FUNCTION_BLOCK FB_StartupReadiness_Tests EXTENDS TcUnit.FB_TestSuite

Power_To_Home_Handoff();
Abort_Cannot_Become_Online();
Error_And_Park_Win();
Completion_Requires_Operational();
Explicit_Abort_Invalidates_Completed_Startup();
Repeated_Start_Does_Not_Reset_Calibration();
Suspended_Automatic_Needs_New_Startup();
Start_While_Initialized_Restarts_Calibration();
Error_Needs_New_Startup();
Parking_Invalidates_Completed_Startup();
Preparation_Stays_0_7_Until_Calibrating();

METHOD PRIVATE Power_To_Home_Handoff
VAR
    fb : BROTLib.FB_StartupReadiness;
END_VAR
TEST('Power_To_Home_Handoff');
fb(Start := TRUE, Parked := TRUE);
AssertEquals_LREAL(0.7, fb.ReadyState, 0.0001, 'preparation, even if parked flag has not cleared');
fb(Start := FALSE, Calibrating := TRUE, Parked := FALSE, Operational := TRUE);
AssertEquals_LREAL(0.8, fb.ReadyState, 0.0001, 'calibration, axes mechanically ready');
fb(Calibrating := FALSE);
AssertEquals_LREAL(0.8, fb.ReadyState, 0.0001, 'handoff/intermediate standstill stays pending');
fb(Completed := TRUE);
AssertEquals_LREAL(1.0, fb.ReadyState, 0.0001, 'only terminal completion is online');
fb(Completed := FALSE);
AssertEquals_LREAL(1.0, fb.ReadyState, 0.0001, 'ordinary subsequent movement remains online');
TEST_FINISHED();
END_METHOD

METHOD PRIVATE Abort_Cannot_Become_Online
VAR
    fb : BROTLib.FB_StartupReadiness;
END_VAR
TEST('Abort_Cannot_Become_Online');
fb(Start := TRUE, Calibrating := TRUE, Operational := TRUE);
fb(Start := FALSE, Aborted := TRUE, Completed := TRUE);
AssertEquals_LREAL(-2.0, fb.ReadyState, 0.0001, 'abort wins over completion');
fb(Aborted := FALSE, Completed := FALSE);
AssertFalse(fb.Initialized, 'enabled axes after abort are not complete');
AssertEquals_LREAL(-2.0, fb.ReadyState, 0.0001, 'clearing flags cannot restore online');
fb(Start := TRUE, Calibrating := FALSE);
AssertEquals_LREAL(0.7, fb.ReadyState, 0.0001, 'retry starts cleanly');
TEST_FINISHED();
END_METHOD

METHOD PRIVATE Error_And_Park_Win
VAR
    fb : BROTLib.FB_StartupReadiness;
END_VAR
TEST('Error_And_Park_Win');
fb(Start := TRUE, Calibrating := TRUE, Completed := TRUE, Operational := TRUE, Error := TRUE);
AssertEquals_LREAL(-1.0, fb.ReadyState, 0.0001, 'error wins');
fb(Start := FALSE, Completed := FALSE, Error := FALSE, Parking := TRUE);
AssertEquals_LREAL(0.3, fb.ReadyState, 0.0001, 'parking');
fb(Parking := FALSE, Parked := TRUE);
AssertEquals_LREAL(0.0, fb.ReadyState, 0.0001, 'parked');
fb(Parked := FALSE);
AssertEquals_LREAL(-2.0, fb.ReadyState, 0.0001, 'no old success after park');
TEST_FINISHED();
END_METHOD

METHOD PRIVATE Completion_Requires_Operational
VAR
    fb : BROTLib.FB_StartupReadiness;
END_VAR
TEST('Completion_Requires_Operational');
fb(Start := TRUE, Calibrating := TRUE, Completed := TRUE, Operational := FALSE);
AssertEquals_LREAL(0.8, fb.ReadyState, 0.0001, 'unfinished focus/not operational prevents completion');
fb(Start := FALSE, Operational := TRUE);
AssertEquals_LREAL(1.0, fb.ReadyState, 0.0001, 'completion with all prerequisites');
fb(Completed := FALSE, Operational := FALSE);
AssertTrue(fb.Initialized, 'transient operational loss preserves completed startup');
AssertEquals_LREAL(-2.0, fb.ReadyState, 0.0001, 'interlock still gates online immediately');
fb(Operational := TRUE);
AssertEquals_LREAL(1.0, fb.ReadyState, 0.0001, 'operational recovery needs no repeated calibration');
TEST_FINISHED();
END_METHOD

METHOD PRIVATE Repeated_Start_Does_Not_Reset_Calibration
VAR
    fb : BROTLib.FB_StartupReadiness;
END_VAR
TEST('Repeated_Start_Does_Not_Reset_Calibration');
fb(Start := TRUE, Calibrating := TRUE, Operational := TRUE);
fb(Calibrating := FALSE);
AssertEquals_LREAL(0.8, fb.ReadyState, 0.0001, 'held/duplicate request does not rewind phase');
fb(Start := FALSE, Completed := TRUE);
AssertTrue(fb.Initialized, 'complete');
fb(Start := TRUE, Completed := FALSE);
AssertEquals_LREAL(0.7, fb.ReadyState, 0.0001, 'accepted new startup clears prior success');
TEST_FINISHED();
END_METHOD

METHOD PRIVATE Explicit_Abort_Invalidates_Completed_Startup
VAR
    fb : BROTLib.FB_StartupReadiness;
END_VAR
TEST('Explicit_Abort_Invalidates_Completed_Startup');
fb(Start := TRUE, Calibrating := TRUE, Completed := TRUE, Operational := TRUE);
AssertTrue(fb.Initialized, 'startup complete');
fb(Start := FALSE, Completed := FALSE, Aborted := TRUE, Operational := FALSE);
AssertFalse(fb.Initialized, 'explicit abort invalidates completed startup');
fb(Aborted := FALSE, Operational := TRUE);
AssertEquals_LREAL(-2.0, fb.ReadyState, 0.0001, 'unlike an interlock, explicit abort needs a new init');
TEST_FINISHED();
END_METHOD

METHOD PRIVATE Suspended_Automatic_Needs_New_Startup
VAR
    fb : BROTLib.FB_StartupReadiness;
END_VAR
TEST('Suspended_Automatic_Needs_New_Startup');
fb(Start := TRUE, Calibrating := TRUE, Completed := TRUE, Operational := TRUE);
AssertEquals_LREAL(1.0, fb.ReadyState, 0.0001, 'online before manual mode');
fb(Start := FALSE, Calibrating := FALSE, Completed := FALSE, Aborted := TRUE, Operational := FALSE);
AssertEquals_LREAL(-2.0, fb.ReadyState, 0.0001, 'manual mode is not online');
fb(Aborted := FALSE, Operational := TRUE);
AssertEquals_LREAL(-2.0, fb.ReadyState, 0.0001, 'back in automatic mode stays offline until a new init');
fb(Start := TRUE);
AssertEquals_LREAL(0.7, fb.ReadyState, 0.0001, 'new init starts again');
TEST_FINISHED();
END_METHOD

METHOD PRIVATE Start_While_Initialized_Restarts_Calibration
VAR
    fb : BROTLib.FB_StartupReadiness;
END_VAR
TEST('Start_While_Initialized_Restarts_Calibration');
fb(Start := TRUE, Calibrating := TRUE, Completed := TRUE, Operational := TRUE);
fb(Start := FALSE, Completed := FALSE, Operational := FALSE);
AssertTrue(fb.Initialized, 'interlock keeps completed startup');
fb(Start := TRUE, Calibrating := FALSE);
AssertFalse(fb.Initialized, 'a Start request discards it, so controllers must not issue one while Initialized');
AssertEquals_LREAL(0.7, fb.ReadyState, 0.0001, 'full startup again');
TEST_FINISHED();
END_METHOD

METHOD PRIVATE Error_Needs_New_Startup
VAR
    fb : BROTLib.FB_StartupReadiness;
END_VAR
TEST('Error_Needs_New_Startup');
fb(Start := TRUE, Calibrating := TRUE, Completed := TRUE, Operational := TRUE);
fb(Start := FALSE, Completed := FALSE, Error := TRUE);
AssertEquals_LREAL(-1.0, fb.ReadyState, 0.0001, 'error');
AssertFalse(fb.Initialized, 'error invalidates completed startup');
fb(Error := FALSE);
AssertEquals_LREAL(-2.0, fb.ReadyState, 0.0001, 'cleared error is not online without a new init');
TEST_FINISHED();
END_METHOD

METHOD PRIVATE Parking_Invalidates_Completed_Startup
VAR
    fb : BROTLib.FB_StartupReadiness;
END_VAR
TEST('Parking_Invalidates_Completed_Startup');
fb(Start := TRUE, Calibrating := TRUE, Completed := TRUE, Operational := TRUE);
fb(Start := FALSE, Completed := FALSE, Parking := TRUE);
AssertEquals_LREAL(0.3, fb.ReadyState, 0.0001, 'parking');
AssertFalse(fb.Initialized, 'parking invalidates completed startup');
fb(Parking := FALSE, Parked := TRUE);
AssertEquals_LREAL(0.0, fb.ReadyState, 0.0001, 'parked');
TEST_FINISHED();
END_METHOD

METHOD PRIVATE Preparation_Stays_0_7_Until_Calibrating
VAR
    fb : BROTLib.FB_StartupReadiness;
END_VAR
TEST('Preparation_Stays_0_7_Until_Calibrating');
fb(Start := TRUE, Operational := TRUE);
AssertEquals_LREAL(0.7, fb.ReadyState, 0.0001, 'preparation');
fb(Start := FALSE);
AssertEquals_LREAL(0.7, fb.ReadyState, 0.0001, 'still preparation without calibration');
fb(Calibrating := TRUE);
AssertEquals_LREAL(0.8, fb.ReadyState, 0.0001, 'calibration');
fb(Calibrating := FALSE);
AssertEquals_LREAL(0.8, fb.ReadyState, 0.0001, 'calibration is not undone by a quiet scan');
TEST_FINISHED();
END_METHOD

END_FUNCTION_BLOCK

(* stored: Version 1.1.0.1, ProductVersion 3.1.4024.15
   POU FB_StartupReadiness_Tests: Id {c2de3b13-6338-437e-a35b-5ebc43113878}, SpecialFunc None
   Method Power_To_Home_Handoff: Id {1b0ac36a-9d5e-4f27-8424-ea7230f7a68f}
   Method Abort_Cannot_Become_Online: Id {6b14a82a-f957-45c4-b97d-8ab02dcec312}
   Method Error_And_Park_Win: Id {7d124066-6035-4ae0-8568-5397f3d2b99f}
   Method Completion_Requires_Operational: Id {3033074d-150f-4719-b3c7-855d2c447217}
   Method Repeated_Start_Does_Not_Reset_Calibration: Id {31b86714-6425-4799-bfe4-559e296f7851}
   Method Explicit_Abort_Invalidates_Completed_Startup: Id {68f3f00d-9ca2-4813-aaac-7e218d1c3586}
   Method Suspended_Automatic_Needs_New_Startup: Id {87b41991-06d0-4e83-842c-e25251082520}
   Method Start_While_Initialized_Restarts_Calibration: Id {73c7d07c-8679-47d5-8fd0-b8dd3b41e731}
   Method Error_Needs_New_Startup: Id {1d95150f-0476-4f8d-a6f3-687167cee33d}
   Method Parking_Invalidates_Completed_Startup: Id {c9fb2c8f-3678-4346-81a7-6fdc609ab8f1}
   Method Preparation_Stays_0_7_Until_Calibrating: Id {ff773175-22de-4aa4-a146-a2152930dec4} *)
